{attribute 'linkalways'}
{attribute 'no_explicit_call' := 'Use the methods of this class'}
{attribute 'enable_dynamic_creation'}
FUNCTION_BLOCK DigitalOut_SimulatedLidarPower IMPLEMENTS I_DigitalOut

METHOD SwitchOn
SimulatorIo.command.isLidarPowered := TRUE;
END_METHOD

METHOD SwitchOff
SimulatorIo.command.isLidarPowered := FALSE;
END_METHOD

PROPERTY IsOn : BOOL
GET
IsOn := SimulatorIo.command.isLidarPowered;
END_GET
END_PROPERTY

END_FUNCTION_BLOCK

(* stored: Version 1.1.0.1, ProductVersion 3.1.4026.12
   POU DigitalOut_SimulatedLidarPower: Id {243003c7-d927-5a12-93fe-9aa1f43afc6f}, SpecialFunc None
   Method SwitchOn: Id {d4eaa0b9-30be-533e-9867-d3301cd5a44b}
   Method SwitchOff: Id {6cced5eb-1e30-5a7f-b154-1c01b9af7853}
   Property IsOn: Id {4f6541ec-7946-5147-82bd-3e6dd9e5f304}
   Get Get: Id {3defebcf-26de-52cb-a7cb-918d176972ca} *)
